# EPICS substitutions: db/Beckhoff_3XXX/ecmcELM3504.substitutions
file "ecmc_analogInputArray-chX.template"
{
  pattern {CH_ID, DTYP,                FTVL  ,  EGU }
          {01,    "asynInt32ArrayIn",  "LONG" , "Raw"}
          {02,    "asynInt32ArrayIn",  "LONG" , "Raw"}
          {03,    "asynInt32ArrayIn",  "LONG" , "Raw"}
          {04,    "asynInt32ArrayIn",  "LONG" , "Raw"}
}

file "ecmcELM360X-stat-chX.template"
{
  pattern {CH_ID}
          {01   }
          {02   }
          {03   }
          {04   }
}

file "ecmc_controlWord-chX.template"
{
  pattern {CH_ID, KEY,   suffix,  sourceName, DESC             }
          {01,    "AI", "-Ctrl", "control",   "AI Control Word"}
          {02,    "AI", "-Ctrl", "control",   "AI Control Word"}
          {03,    "AI", "-Ctrl", "control",   "AI Control Word"}
          {04,    "AI", "-Ctrl", "control",   "AI Control Word"}
}
